{attribute 'linkalways'} 
{attribute 'no_explicit_call' := 'This FB is a CLASS and must be accessed using methods or properties'}
{attribute 'enable_dynamic_creation'}
FUNCTION_BLOCK Mc2AxisSoeDrive EXTENDS Mc2Axis IMPLEMENTS Axis, Drive
VAR
	reset_drive_command2 : ResetSoeDriveCommand(axis := THIS^);
END_VAR

METHOD PUBLIC CyclicCall
SUPER^.CyclicCall();

reset_drive_command.CyclicCall();
END_METHOD

METHOD PUBLIC ResetDrive : AsyncCommand
reset_drive_command2.Execute();
ResetDrive := reset_drive_command2;
END_METHOD

END_FUNCTION_BLOCK

(* stored: Version 1.1.0.1
   POU Mc2AxisSoeDrive: Id {f9336e12-837f-4479-a744-0cde172ef32e}, SpecialFunc None
   Folder Administrative: Id {a31e2a5d-92ba-4dbc-a584-749921522786}
   Folder Cyclic: Id {2a8a0a3a-db02-4f79-9dd6-f81e7b90e64e}
   Folder Properties: Id {d0057c44-c327-4610-8a8f-f1ef5d4b11f5}
   Folder Error: Id {ab1d5148-4ec5-43f8-ac28-278a9506a8ff}
   Method CyclicCall: Id {4b3d7009-6e56-41f2-b11e-2d69af3fb445}
   Method ResetDrive: Id {9280250d-0d91-4024-9e78-cfb30ab3c1b5} *)
